// TIA Portal project "AT2_Start_Uebung" (V18)

(* hardware
DEVICE "PLC_1_Station"  S7-1500 station
   slot 0: "Profilschiene_0"  Rack  6ES7 590-1***0-0AA0
   slot 1: "PLC_1"  CPU 1516-3 PN/DP  6ES7 516-3AN02-0AB0  V2.8
      slot 3: "CPU-Display_1"  6ES7591-1BA00-0AA0
      slot 32768: "PROFINET-Schnittstelle_1"  X1
         slot 32769: "Port_1"  X1 P1
         slot 32770: "Port_2"  X1 P2
      slot 33024: "PROFINET-Schnittstelle_2"  X2
         slot 33025: "Port_1"  X2 P1
      slot 33280: "DP-Schnittstelle_1"  X3
      slot 34817: "Virtual CP interface port_1"  Virtual CP interface port  Virtual CP interface port
*)

// ===== PLC "PLC_1"  CPU 1516-3 PN/DP =====

VAR_GLOBAL   // PLC tag table "AT2_Vorgegebene_Merker"
   "DAUER EIN" AT %M0.1 : Bool;   // Vorgegebener Merker aus AT-2 Anhang S. 2.
   "Freigabe Messung" AT %M2.5 : Bool;   // Vorgegebener Merker aus AT-2 Anhang S. 2.
   "Test Messung EIN" AT %M4.0 : Bool;   // Vorgegebener Merker aus AT-2 Anhang S. 2.
   "Test Messung Links fahren" AT %M4.1 : Bool;   // Vorgegebener Merker aus AT-2 Anhang S. 2.
   "Test Messung Rechts fahren" AT %M4.2 : Bool;   // Vorgegebener Merker aus AT-2 Anhang S. 2.
   "Impulse Test Messung" AT %MD20 : DInt;   // Anhang S. 2; numerische Adressen entzerrt, siehe STARTZUSTAND.md.
   "Impulse Zurücksetzen" AT %M4.3 : Bool;   // Vorgegebener Merker aus AT-2 Anhang S. 2.
   "Impulse Längenmessung" AT %MD24 : DInt;   // Anhang S. 2; numerische Adressen entzerrt, siehe STARTZUSTAND.md.
   "Länge in mm" AT %M10.0 : LReal;   // Anhang S. 2; numerische Adressen entzerrt, siehe STARTZUSTAND.md.
END_VAR

DATA_BLOCK "IEC_Counter_0_DB"   // DB2
{ S7_Optimized_Access := 'TRUE' }
AUTHOR : SIMATIC
FAMILY : IEC
NAME : DCNTR
VERSION : 1.2
// stored: InstanceOfName IEC_DCOUNTER
"IEC_DCOUNTER"
BEGIN
END_DATA_BLOCK

FUNCTION "1_Geschwindigkeitsvorwahl" : Void   // FC1, FBD
{ S7_Optimized_Access := 'TRUE' }
// Rekonstruierter Übungsstart, keine originale Hochschul-Projektdatei.
   VAR_INPUT
      Aktivierung : Bool;
      "Geschwindigkeitsvorgabe in % IN" : Real;
   END_VAR
   VAR_TEMP
      "Fehler Scale TEMP" : Word;
      Temp : Int;
   END_VAR
BEGIN

REGION Network 1: Geschwindigkeitsvorwahl
   // Vorgegebener UNSCALE-Aufruf aus Anhang S. 6. Ausgangszuordnung und Geschwindigkeitswahl bleiben Übungsaufgaben.
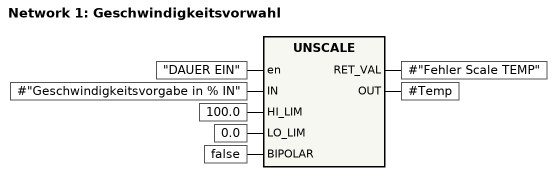
   IF "DAUER EIN" THEN
       #"Fehler Scale TEMP" := UNSCALE(IN := #"Geschwindigkeitsvorgabe in % IN",
                               HI_LIM := 100.0,
                               LO_LIM := 0.0,
                               BIPOLAR := false,
                               OUT => #Temp);
   END_IF;
END_REGION
END_FUNCTION

FUNCTION "2_Ansteuerung Motor" : Void   // FC2, FBD
{ S7_Optimized_Access := 'TRUE' }
// Rekonstruierter Übungsstart, keine originale Hochschul-Projektdatei.
   VAR_INPUT
      "Band nach links fahren EIN" : Bool;
      "Band nach rechts fahren EIN" : Bool;
   END_VAR
BEGIN

REGION Network 1: Motoransteuerung Band rechts
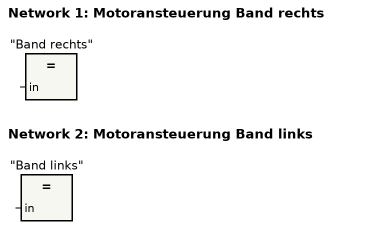
   "Band rechts" := TRUE;
END_REGION

REGION Network 2: Motoransteuerung Band links
   "Band links" := TRUE;
END_REGION
END_FUNCTION

FUNCTION "Längenmessung" : Void   // FC3, FBD
{ S7_Optimized_Access := 'TRUE' }
// Rekonstruierter Übungsstart, keine originale Hochschul-Projektdatei.
BEGIN

REGION Network 1: Längenmessung
   // AT-2 Aufgabe 2.2: Schnittstelle und Messfunktion selbst erstellen. Im Anhang ist keine fertige FC3-Schaltung abgebildet.
END_REGION
END_FUNCTION

FUNCTION "6_Test Messung" : Void   // FC6, FBD
{ S7_Optimized_Access := 'TRUE' }
// Rekonstruierter Übungsstart, keine originale Hochschul-Projektdatei.
   VAR_INPUT
      "Rücksetzen der Impulse" : Bool;
   END_VAR
   VAR_OUTPUT
      Impulse : DInt;
   END_VAR
BEGIN

REGION Network 1: Test Messung
   // Vorgegebener Prüfbaustein aus Anhang S. 5. Fehlende I/O-Symbole und Motorzustände selbst zuordnen.
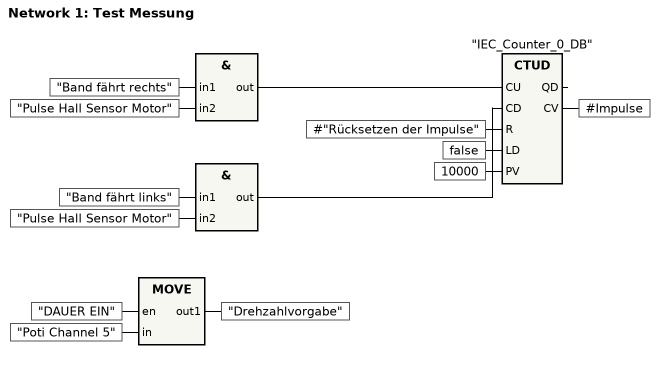
   "IEC_Counter_0_DB".CTUD(CU := "Band fährt rechts" AND "Pulse Hall Sensor Motor",
                           CD := "Band fährt links" AND "Pulse Hall Sensor Motor",
                           R := #"Rücksetzen der Impulse",
                           LD := false,
                           PV := 10000,
                           CV => #Impulse);
   IF "DAUER EIN" THEN "Drehzahlvorgabe" := "Poti Channel 5"; END_IF;
END_REGION
END_FUNCTION

ORGANIZATION_BLOCK "Main"   // OB1, FBD, ProgramCycle
TITLE = "Main Program Sweep (Cycle)"
{ S7_Optimized_Access := 'TRUE' }
VERSION : 0.1
// Rekonstruierter Übungsstart, keine originale Hochschul-Projektdatei.
   VAR_INPUT
      Initial_Call : Bool;   // Initial call of this OB
      Remanence : Bool;   // =True, if remanent data are available
   END_VAR
BEGIN

REGION Network 1: DAUER EIN
END_REGION

REGION Network 2: Ansteuerung Motor
END_REGION

REGION Network 3: Test Messung
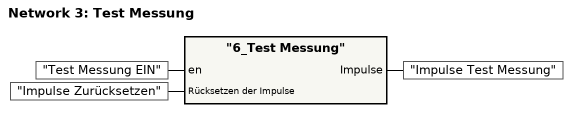
   IF "Test Messung EIN" THEN
       "6_Test Messung"("Rücksetzen der Impulse" := "Impulse Zurücksetzen", Impulse => "Impulse Test Messung");
   END_IF;
END_REGION

REGION Network 4: Längenmessung
END_REGION

REGION Network 5: Freigabe Messung
END_REGION
END_ORGANIZATION_BLOCK